VISUALIZATION FP_Drive  // 1024x768
END_VISUALIZATION

(* stored: Version 1.1.0.1
   Visu FP_Drive: Id {78112fab-05fc-4177-a21e-7580a845d322} *)
